(* IEC 61131-3 sources: plcassist-cli/packages/volt-lsp-iec/test-corpus/bakon-nano/Device/Plc Logic/Application/Library Manager/CmpAsyncMgr, 10 files *)

(* ---- GVL.gvl ---- *)
VAR_GLOBAL
	ASYNCJOB_INVALID_HANDLE : RTS_IEC_HANDLE := RTS_INVALID_HANDLE;
	ASYNCJOB_TASK : UDINT := 0;
	ASYNCJOB_EVENT : UDINT := 1;
	ASYNCJOB_HOOK : UDINT := 2;
	ASYNCSTATE_INVALID : UDINT := 16#FFFFFFFF;
	ASYNCSTATE_PENDING : UDINT := 0;
	ASYNCSTATE_ACTIVE : UDINT := 1;
	ASYNCSTATE_READY : UDINT := 2;
	ASYNCSTATE_ERROR : UDINT := 3;
	ASYNCSTATE_TIMEOUT : UDINT := 4;
	ASYNC_TIMEOUT_INFINITE : UDINT := 0;
	ASYNC_IS_IEC : UDINT := 1;
	ASYNC_ISNOT_IEC : UDINT := 0;
	CH_COMM_CYCLE : UDINT := 20;
END_VAR

(* ---- GVL_2.gvl ---- *)
VAR_GLOBAL
	CMPASYNCMGR_VERSION_3_5_6_0 : BOOL := TRUE;
END_VAR

(* ---- TASK_PRIORITIES.gvl ---- *)
VAR_GLOBAL
	TASKPRIO_RANGE : UDINT := 255;
	TASKPRIO_SEGMENT : UDINT := 32;
	TASKPRIO_MAX : UDINT := 0;
	TASKPRIO_SYSTEM_BASE : UDINT := 0;
	TASKPRIO_SYSTEM_END : UDINT := 31;
	TASKPRIO_REALTIME_BASE : UDINT := 32;
	TASKPRIO_REALTIME_END : UDINT := 63;
	TASKPRIO_HIGH_BASE : UDINT := 64;
	TASKPRIO_HIGH_END : UDINT := 95;
	TASKPRIO_ABOVENORMAL_BASE : UDINT := 96;
	TASKPRIO_ABOVENORMAL_END : UDINT := 127;
	TASKPRIO_NORMAL_BASE : UDINT := 128;
	TASKPRIO_NORMAL_END : UDINT := 159;
	TASKPRIO_BELOWNORMAL_BASE : UDINT := 160;
	TASKPRIO_BELOWNORMAL_END : UDINT := 191;
	TASKPRIO_LOW_BASE : UDINT := 192;
	TASKPRIO_LOW_END : UDINT := 223;
	TASKPRIO_LOWEST_BASE : UDINT := 224;
	TASKPRIO_LOWEST_END : UDINT := 255;
	TASKPRIO_IDLE : UDINT := 255;
	TASKPRIO_MIN : UDINT := 255;
END_VAR

(* ---- ASYNCADD.fun ---- *)
FUNCTION ASYNCADD : RTS_IEC_HANDLE
VAR_INPUT
	PFJOBFUNC : POINTER TO BYTE;
	PPARAM : POINTER TO BYTE;
	PINSTANCE : POINTER TO BYTE;
	PULSTATE : POINTER TO UDINT;
	ULIECFUNC : UDINT;
	ULTYPE : UDINT;
	ULTIMEOUT : UDINT;
	PASYNCJOBPARAM : POINTER TO ASYNCJOB_PARAM;
	PRESULT : POINTER TO RTS_IEC_RESULT;
END_VAR
END_FUNCTION

(* ---- ASYNCGETJOBRETURNVALUE.fun ---- *)
FUNCTION ASYNCGETJOBRETURNVALUE : RTS_IEC_RESULT
VAR_INPUT
	HJOB : RTS_IEC_HANDLE;
	PULRETURNVAL : POINTER TO UDINT;
END_VAR
END_FUNCTION

(* ---- ASYNCGETNUMOFJOBS.fun ---- *)
FUNCTION ASYNCGETNUMOFJOBS : RTS_IEC_RESULT
VAR_IN_OUT
	NUMOFJOBS : ASYNCJOB_CURRENT_MAX;
	NUMOFJOBTASKS : ASYNCJOB_CURRENT_MAX;
END_VAR
END_FUNCTION

(* ---- ASYNCKILL.fun ---- *)
FUNCTION ASYNCKILL : RTS_IEC_RESULT
VAR_INPUT
	HJOB : RTS_IEC_HANDLE;
END_VAR
END_FUNCTION

(* ---- ASYNCREMOVE.fun ---- *)
FUNCTION ASYNCREMOVE : RTS_IEC_RESULT
VAR_INPUT
	HJOB : RTS_IEC_HANDLE;
END_VAR
END_FUNCTION

(* ---- ASYNCREMOVEALL.fun ---- *)
FUNCTION ASYNCREMOVEALL : RTS_IEC_RESULT
END_FUNCTION

(* ---- ASYNCBASECLASS.fb ---- *)
FUNCTION_BLOCK ASYNCBASECLASS
VAR
	ULTYPE : UDINT;
	ULTOUT : UDINT;
	PJOBPARAMS : POINTER TO ASYNCJOB_PARAM;
END_VAR
END_FUNCTION_BLOCK

METHOD ASYNCREMOVEJOB : RTS_IEC_RESULT
VAR_INPUT
	HJOB : RTS_IEC_HANDLE;
END_VAR
END_METHOD

METHOD ASYNCSETJOBPARAMS : RTS_IEC_RESULT
VAR_INPUT
	ULASYNCJOBTYPE : UDINT;
	ULTIMEOUT : UDINT;
	PASYNCJOBPARAMS : POINTER TO ASYNCJOB_PARAM;
END_VAR
END_METHOD
